{region 'Documentation'}
(*!
<summary>Check that IN is inside the inclusive StartTime..EndTime interval.</summary>
<description>

StartTime &gt; EndTime reports Error during active evaluation; equal bounds are
valid.

Compares calendar days only; hidden time-of-day components are ignored.

</description>
*)
{endregion}
FUNCTION_BLOCK AssertInTimespan_Date EXTENDS AssertionBase
VAR_INPUT
    IN : DATE; //! Actual value checked or observed by this Assertion.
    StartTime : DATE; //! Inclusive start of the time span; must not exceed EndTime.
    EndTime : DATE; //! Inclusive end of the time span; must not precede StartTime.
END_VAR

SUPER^();

{region 'Documentation'}
(*!
<summary>Evaluate the typed temporal relation and report higher-priority errors first.</summary>
*)
{endregion}
METHOD PROTECTED Assert
VAR
    Message : STRING(GVL_Constants.MessageLength);
    StartTimeText : STRING(GVL_Constants.AssertionValueLength);
    EndTimeText : STRING(GVL_Constants.AssertionValueLength);
    ActualText : STRING(GVL_Constants.AssertionValueLength);
END_VAR
IF NOT EvaluationActive THEN
    RETURN;
END_IF;

IF Result = E_Result.Error THEN
    RETURN;
END_IF;

IF DateToDayNumber(Value := StartTime) > DateToDayNumber(Value := EndTime) THEN
    StartTimeText := DATE_TO_STRING(StartTime);
    EndTimeText := DATE_TO_STRING(EndTime);
    Message := CONCAT('Assertion error: start time exceeds end time. StartTime = ',
        StartTimeText);
    Message := CONCAT(Message, ', EndTime = ');
    Message := CONCAT(Message, EndTimeText);
    Message := CONCAT(Message, '.');
    Error(Message := Message);
    RETURN;
END_IF;

IF Result = E_Result.Failed THEN
    RETURN;
END_IF;

IF (DateToDayNumber(Value := IN) < DateToDayNumber(Value := StartTime))
    OR (DateToDayNumber(Value := IN) > DateToDayNumber(Value := EndTime)) THEN
    StartTimeText := DATE_TO_STRING(StartTime);
    EndTimeText := DATE_TO_STRING(EndTime);
    ActualText := DATE_TO_STRING(IN);
    Message := CONCAT('Assertion failed: value is outside allowed timespan. StartTime = ',
        StartTimeText);
    Message := CONCAT(Message, ', EndTime = ');
    Message := CONCAT(Message, EndTimeText);
    Message := CONCAT(Message, ', Actual = ');
    Message := CONCAT(Message, ActualText);
    Message := CONCAT(Message, '.');
    Fail(Message := Message);
    RETURN;
END_IF;

Pass();
END_METHOD

END_FUNCTION_BLOCK

(* stored: Version 1.1.0.1
   POU AssertInTimespan_Date: Id {24c1958d-a258-4649-af18-a387360c4dcf}, SpecialFunc None
   Folder Internal: Id {aa226307-1024-42cc-9adb-bd341656a66a}
   Method Assert: Id {76112a32-49bb-425b-b38c-644b879c0ef9} *)
